{region 'Documentation'}
(*!
<summary>Check that IN is greater than Minimum.</summary>
*)
{endregion}
FUNCTION_BLOCK AssertGreaterThan_SInt EXTENDS AssertionBase
VAR_INPUT
    IN : SINT; //! Actual value checked or observed by this Assertion.
    Minimum : SINT; //! Exclusive lower bound; the actual value or count must be greater.
END_VAR

SUPER^();

{region 'Documentation'}
(*!
<summary>Check that IN is greater than Minimum.</summary>
*)
{endregion}
METHOD PROTECTED Assert
VAR
    Message : STRING(GVL_Constants.MessageLength);
    MinimumText : STRING(GVL_Constants.AssertionValueLength);
    ActualText : STRING(GVL_Constants.AssertionValueLength);
END_VAR
IF NOT EvaluationActive THEN
    RETURN;
END_IF;

IF Result = E_Result.Error THEN
    RETURN;
END_IF;

IF Result = E_Result.Failed THEN
    RETURN;
END_IF;

IF IN <= Minimum THEN
    MinimumText := SINT_TO_STRING(Minimum);
    ActualText := SINT_TO_STRING(IN);
    Message := CONCAT('Assertion failed: value is not greater than minimum. Minimum = ',
        MinimumText);
    Message := CONCAT(Message, ', Actual = ');
    Message := CONCAT(Message, ActualText);
    Message := CONCAT(Message, '.');
    Fail(Message := Message);
    RETURN;
END_IF;

Pass();
END_METHOD

END_FUNCTION_BLOCK

(* stored: Version 1.1.0.1
   POU AssertGreaterThan_SInt: Id {b4b9600d-18a1-482c-9fb3-56ec8f23b47f}, SpecialFunc None
   Folder Internal: Id {f9a1370a-e284-4036-aa0a-eb2b7ac380b3}
   Method Assert: Id {affa6a3c-359e-48d5-b9a0-874deb6e9dab} *)
